(* IEC 61131-3 sources: veristc/veri-ide/tests/fixtures/valid-project/logic, 2 files *)

(* ---- pid.st ---- *)
FUNCTION_BLOCK pid
VAR_INPUT
    setpoint : DINT;
    process_value : DINT;
END_VAR

VAR_OUTPUT
    control_output : DINT;
END_VAR

VAR
    error : DINT;
    kp : DINT := 10;
END_VAR

error := setpoint - process_value;
control_output := error * kp;

END_FUNCTION_BLOCK

(* ---- MAIN.st ---- *)
PROGRAM main
VAR
    counter : DINT;
    status : DINT;
END_VAR

counter := counter + 1;
IF counter > 100 THEN
    counter := 0;
    status := 1;
END_IF;

END_PROGRAM
